(* PLC project HeatExchanger_PLC_Control.project, CODESYS CODESYS V3.5 SP22 Patch 4 *)
(* stored: creationDateTime 2026-10-29T16:53:11.6519631, modificationDateTime 2026-10-29T16:50:30.2076377 *)

PROGRAM PLC_PRG
  VAR
    plant : FB_PlantSim;
    ctrl : FB_TempControl;
    sp : REAL := 0.0;  (* temperature setpoint, degC rise *)
    useSmith : BOOL := FALSE;  (* FALSE = PI, TRUE = PI with Smith predictor *)
    manualMode : BOOL := FALSE;  (* TRUE = operator sets the valve *)
    manualOut : REAL := 0.0;  (* operator valve position, % *)
    filterOn : BOOL := FALSE;  (* measurement filter *)
    noiseOn : BOOL := FALSE;  (* sensor noise *)
    dist : REAL := 0.0;  (* input disturbance, % valve *)
    gainFactor : REAL := 1.0;  (* plant gain change (1.3 or 0.7) *)
    delayFactor : REAL := 1.0;  (* plant delay change (1.3 or 0.7) *)
    temp : REAL;  (* measured temperature rise, degC *)
    valve : REAL;  (* valve command, % *)
    alarm : FB_Alarm;  (* alarms and interlock *)
    ackBtn : BOOL;  (* operator acknowledge *)
    resetBtn : BOOL;  (* operator interlock reset *)
  END_VAR

                    // alarms: check the measurement first
alarm(pv := plant.y, ack := ackBtn, reset := resetBtn);

// controller: reads the measurement from the previous scan
// interlock forces manual mode with the valve closed (0 %)
ctrl(sp := sp, pv := plant.y, useSmith := useSmith,
     manualMode := manualMode OR alarm.interlock,
     manualOut  := SEL(alarm.interlock, manualOut, 0.0),
     filterOn := filterOn);
valve := ctrl.u;

// simulated heat exchanger
plant(u := valve, dist := dist, gainFactor := gainFactor,
      delayFactor := delayFactor, noiseOn := noiseOn);
temp := plant.y;
                  
END_PROGRAM

FUNCTION_BLOCK FB_PlantSim
  VAR_INPUT
    u : REAL;  (* heating valve position, % *)
    dist : REAL;  (* input disturbance, % valve *)
    gainFactor : REAL := 1.0;  (* 1.3 or 0.7 for the robustness cases *)
    delayFactor : REAL := 1.0;  (* 1.3 or 0.7 for the robustness cases *)
    noiseOn : BOOL;
  END_VAR
  VAR_OUTPUT
    y : REAL;  (* measured temperature rise, degC *)
    yClean : REAL;  (* measured value without noise *)
  END_VAR
  VAR
    K : REAL := 1.5;  (* gain, degC per % valve *)
    tau : REAL := 50.0;  (* time constant, s *)
    theta : REAL := 15.0;  (* transport delay, s *)
    tauS : REAL := 5.0;  (* sensor lag, s *)
    Ts : REAL := 0.1;  (* scan time, s *)
    buf : ARRAY[0..399] OF REAL;
    wr : INT := 0;
    rd : INT;
    nd : INT;
    ud : REAL;
    x : REAL;
    ys : REAL;
    alpha : REAL;
    beta : REAL;
    seed : DWORD := 12345;
    i : INT;
    sumU : REAL;
  END_VAR

                    alpha := EXP(-Ts / tau);
beta  := EXP(-Ts / tauS);

// delay in samples, limited to the buffer size
nd := REAL_TO_INT(theta * delayFactor / Ts);
IF nd < 0 THEN nd := 0; END_IF
IF nd > 399 THEN nd := 399; END_IF

// delay buffer: store the new input, read the old one
buf[wr] := u + dist;
rd := wr - nd;
IF rd < 0 THEN rd := rd + 400; END_IF
ud := buf[rd];
wr := wr + 1;
IF wr > 399 THEN wr := 0; END_IF

// plant lag and sensor lag
x  := alpha * x  + (1.0 - alpha) * K * gainFactor * ud;
ys := beta  * ys + (1.0 - beta)  * x;
yClean := ys;

// measurement noise, about 0.05 degC standard deviation
sumU := 0.0;
FOR i := 1 TO 12 DO
    seed := seed * DWORD#1664525 + DWORD#1013904223;
    sumU := sumU + DWORD_TO_REAL(seed) / 4294967296.0;
END_FOR
IF noiseOn THEN
    y := ys + 0.05 * (sumU - 6.0);
ELSE
    y := ys;
END_IF
                  
END_FUNCTION_BLOCK

FUNCTION_BLOCK FB_PI
  VAR_INPUT
    err : REAL;  (* error = setpoint - measurement (corrected for Smith predictor) *)
    Kc : REAL;  (* controller gain, % valve per degC *)
    Ti : REAL := 50.0;  (* integral time, s *)
    outMin : REAL := 0.0;  (* output low limit, % *)
    outMax : REAL := 100.0;  (* output high limit, % *)
    manual : BOOL;  (* TRUE = manual mode (controller follows manualOut) *)
    manualOut : REAL;  (* valve position set by the operator, % *)
  END_VAR
  VAR_OUTPUT
    u : REAL;  (* valve command, % *)
  END_VAR
  VAR
    Ts : REAL := 0.1;  (* scan time, s *)
    pTerm : REAL;
    intg : REAL;  (* integral term *)
    intgNew : REAL;
    uCand : REAL;
  END_VAR

                    pTerm := Kc * err;

IF manual THEN
    // follow the operator value, so switching back to auto causes no jump
    intg := manualOut - pTerm;
    u := LIMIT(outMin, manualOut, outMax);
ELSE
    IF Ti > 0.001 THEN
        intgNew := intg + Kc * err * Ts / Ti;
    ELSE
        intgNew := intg;
    END_IF
    uCand := pTerm + intgNew;

    // anti-windup: stop integrating while the output is saturated
    // and the error would push it further into the limit
    IF (uCand > outMax AND err > 0.0) OR (uCand < outMin AND err < 0.0) THEN
        ;
    ELSE
        intg := intgNew;
    END_IF
    u := LIMIT(outMin, pTerm + intg, outMax);
END_IF
                  
END_FUNCTION_BLOCK

FUNCTION_BLOCK FB_SmithPredictor
  VAR_INPUT
    u : REAL;  (* controller output (valve command), % *)
    K : REAL := 1.5;  (* model gain, degC per % valve *)
    tau : REAL := 50.0;  (* model time constant, s *)
    theta : REAL := 15.0;  (* model delay, s *)
    tauS : REAL := 5.0;  (* sensor lag in the model, s *)
  END_VAR
  VAR_OUTPUT
    ym0 : REAL;  (* model output without delay *)
    ym : REAL;  (* model output with delay *)
    corr : REAL;  (* correction = ym0 - ym *)
  END_VAR
  VAR
    Ts : REAL := 0.1;  (* scan time, s *)
    buf : ARRAY[0..399] OF REAL;
    wr : INT := 0;
    rd : INT;
    nd : INT;
    ud : REAL;
    x0 : REAL;
    x1 : REAL;
    ys0 : REAL;
    ys1 : REAL;
    alpha : REAL;
    beta : REAL;
  END_VAR

                    alpha := EXP(-Ts / tau);
beta  := EXP(-Ts / tauS);

// model delay in samples
nd := REAL_TO_INT(theta / Ts);
IF nd < 0 THEN nd := 0; END_IF
IF nd > 399 THEN nd := 399; END_IF

// delay buffer for the model with delay
buf[wr] := u;
rd := wr - nd;
IF rd < 0 THEN rd := rd + 400; END_IF
ud := buf[rd];
wr := wr + 1;
IF wr > 399 THEN wr := 0; END_IF

// model without delay: plant lag, then sensor lag
x0  := alpha * x0  + (1.0 - alpha) * K * u;
ys0 := beta  * ys0 + (1.0 - beta)  * x0;

// model with delay: same, but fed with the delayed input
x1  := alpha * x1  + (1.0 - alpha) * K * ud;
ys1 := beta  * ys1 + (1.0 - beta)  * x1;

ym0  := ys0;
ym   := ys1;
corr := ym0 - ym;
                  
END_FUNCTION_BLOCK

FUNCTION_BLOCK FB_TempControl
  VAR_INPUT
    sp : REAL;  (* temperature setpoint, degC rise *)
    pv : REAL;  (* measured temperature, degC rise *)
    useSmith : BOOL;  (* FALSE = PI, TRUE = PI with Smith predictor *)
    manualMode : BOOL;  (* TRUE = operator sets the valve *)
    manualOut : REAL;  (* operator valve position, % *)
    filterOn : BOOL;  (* measurement filter on or off *)
    Tf : REAL := 2.0;  (* filter time constant, s *)
    KcPI : REAL := 0.834;  (* PI tuning (MATLAB final design) *)
    TiPI : REAL := 50.0;
    KcSM : REAL := 3.336;  (* PI tuning used with the Smith predictor *)
    TiSM : REAL := 50.0;
  END_VAR
  VAR_OUTPUT
    u : REAL;  (* heating valve command, % *)
    pvF : REAL;  (* temperature used by the controller *)
    corr : REAL;  (* Smith predictor correction *)
  END_VAR
  VAR
    Ts : REAL := 0.1;  (* scan time, s *)
    piPlain : FB_PI;
    piSmith : FB_PI;
    smith : FB_SmithPredictor;
    errPI : REAL;
    errSM : REAL;
    mo : REAL;
    uPrev : REAL;
  END_VAR

                    // measurement filter (first order), can be switched off
IF filterOn AND (Tf > 0.0) THEN
    pvF := pvF + Ts / (Tf + Ts) * (pv - pvF);
ELSE
    pvF := pv;
END_IF

// errors for the two controllers
errPI := sp - pvF;
errSM := sp - pvF - smith.corr;   // correction from the previous scan

// value the idle controller follows (keeps switching bumpless)
IF manualMode THEN
    mo := manualOut;
ELSE
    mo := uPrev;
END_IF

piPlain(err := errPI, Kc := KcPI, Ti := TiPI,
        manual := (manualMode OR useSmith), manualOut := mo);
piSmith(err := errSM, Kc := KcSM, Ti := TiSM,
        manual := (manualMode OR NOT useSmith), manualOut := mo);

// select the output
IF manualMode THEN
    u := LIMIT(0.0, manualOut, 100.0);
ELSIF useSmith THEN
    u := piSmith.u;
ELSE
    u := piPlain.u;
END_IF
uPrev := u;

// run the predictor models with the new valve command
smith(u := u);
corr := smith.corr;
                  
END_FUNCTION_BLOCK

FUNCTION_BLOCK FB_Alarm
  VAR_INPUT
    pv : REAL;
    ack : BOOL;
    reset : BOOL;
    tahLimit : REAL := 15.0;
    tahhLimit : REAL := 20.0;
    deadband : REAL := 0.5;
  END_VAR
  VAR_OUTPUT
    high : BOOL;
    highHigh : BOOL;
    sensorFault : BOOL;
    interlock : BOOL;
    horn : BOOL;
    state : INT;
  END_VAR
  VAR
    tonH : TON;
    tonHH : TON;
    rtAck : R_TRIG;
    rtReset : R_TRIG;
    rtH : R_TRIG;
    rtHH : R_TRIG;
    rtSF : R_TRIG;
    condH : BOOL;
    condHH : BOOL;
    anyActive : BOOL;
    unacked : BOOL;
  END_VAR

                    IF high THEN condH := pv > (tahLimit - deadband);
ELSE condH := pv > tahLimit; END_IF
tonH(IN := condH, PT := T#2S);
high := tonH.Q;

IF highHigh THEN condHH := pv > (tahhLimit - deadband);
ELSE condHH := pv > tahhLimit; END_IF
tonHH(IN := condHH, PT := T#2S);
highHigh := tonHH.Q;

sensorFault := (pv < -5.0) OR (pv > 60.0);

anyActive := high OR highHigh OR sensorFault;
   rtH(CLK := high);
   rtHH(CLK := highHigh);
   rtSF(CLK := sensorFault);
rtAck(CLK := ack);
rtReset(CLK := reset);

IF rtH.Q OR rtHH.Q OR rtSF.Q THEN unacked := TRUE; END_IF
IF rtAck.Q THEN unacked := FALSE; END_IF
horn := unacked;

IF anyActive THEN
    IF unacked THEN state := 1; ELSE state := 2; END_IF
ELSE
    IF unacked THEN state := 3; ELSE state := 0; END_IF
END_IF

IF highHigh OR sensorFault THEN interlock := TRUE; END_IF
IF rtReset.Q AND NOT highHigh AND NOT sensorFault AND (pv < tahLimit) THEN
    interlock := FALSE;
END_IF
                  
END_FUNCTION_BLOCK

CONFIGURATION Device
  RESOURCE Application ON PLC
    TASK MainTask(INTERVAL := T#100ms, PRIORITY := 1);
    TASK VISU_TASK(INTERVAL := T#100ms, PRIORITY := 31);
    PROGRAM PLC_PRG WITH MainTask : PLC_PRG;
    PROGRAM VisuElems.Visu_Prg WITH VISU_TASK : VisuElems.Visu_Prg;
  END_RESOURCE
END_CONFIGURATION
